(* IEC 61131-3 sources: Lasal-MCP/examples/SampleSource/LASALScreenAdvancedSolution/LASALScreenAdvancedSolution/LASALScreenAdvacnedSolution/Stations/Terminal/HMI/Class/MyRecalculate, 1 file *)

(* ---- MyRecalculate.st ---- *)
(*!
<Class
	Name               = "MyRecalculate"
	Revision           = "0.0"
	RealtimeTask       = "false"
	CyclicTask         = "false"
	BackgroundTask     = "false"
	Sigmatek           = "false"
	OSInterface        = "false"
	HighPriority       = "false"
	Automatic          = "false"
	UpdateMode         = "Prescan"
	SharedCommandTable = "true"
	Objectsize         = "(390,120)">
	<Channels>
		<Server Name="Length" Visualized="true" Initialize="false" WriteProtected="false" Retentive="false"/>
	</Channels>
	<Network Name="MyRecalculate">
		<!-- List of Components in this network -->
		<Components>
			<Object
				Name       = "_base"
				Class      = "_Global"
				Position   = "(218,120)"
				Visualized = "true"
				Remotely   = "true">
				<Channels>
					<Server Name="Server0"/>
					<Client Name="Lse"/>
				</Channels>
			</Object>
		</Components>
		<Comments>
		</Comments>
		<!-- List of Connections in this network -->
		<Connections>
			<Connection Source="this.Server0" Destination="_base.Server0" Vertices="(690,210),(518,210),"/>
			<Connection Source="_base.Lse" Destination="this.Lse" Vertices="(218,210),(38,210),"/>
		</Connections>
		<!-- Headerfiles -->
		<Options>
		</Options>
	</Network>
</Class>
*)
#pragma using _Global

MyRecalculate : CLASS
: _Global
  //Servers:
	Length 	: SvrCh_REAL;
  //Clients:
  //Variables:
  //Functions:
				//! <Function Comment="function is called in case of an recalculation (formula) defined for a data-server&#13;&#10;pres ....... --&gt; to value&#13;&#10;pv ......... --&gt; to variable&#13;&#10;direction .. direction (TRUE Y=kX+d, FALSE X=(Y+d)/k)&#13;&#10;retcode .... return TRUE if kernel should do the calculation, on the other hand return FALSE&#13;&#10;" Name="IF_Recalculate"/>
	FUNCTION VIRTUAL GLOBAL IF_Recalculate
		VAR_INPUT
			pres 	: ^_RESULT;
			pv 	: ^_VARIABLE;
			direction 	: BOOL;
		END_VAR
		VAR_OUTPUT
			retcode 	: BOOL;
		END_VAR;

	FUNCTION MeterToFeet
		VAR_INPUT
			value 	: REAL;
			dir 	: BOOL;
		END_VAR
		VAR_OUTPUT
			retcode 	: REAL;
		END_VAR;
  //Tables:
	FUNCTION @STD
		VAR_OUTPUT
			ret_code	: CONFSTATES;
		END_VAR;
	FUNCTION GLOBAL TAB @CT_;
END_CLASS;

FUNCTION VIRTUAL GLOBAL MyRecalculate::IF_Recalculate
	VAR_INPUT
		pres 	: ^_RESULT;
		pv 	: ^_VARIABLE;
		direction 	: BOOL;
	END_VAR
	VAR_OUTPUT
		retcode 	: BOOL;
	END_VAR

  retcode := TRUE;

  //====================================================================================
  case pv^.info.formula of

    //----------------------------------------------------------------------------------
    50: // The Formula number to be used for the unit

        pres^.value$REAL := MeterToFeet(value:= pres^.value$REAL, dir:= direction);

        retcode := FALSE;

  end_case;

END_FUNCTION

FUNCTION MyRecalculate::MeterToFeet
	VAR_INPUT
		value 	: REAL;
		dir 	: BOOL;
	END_VAR
	VAR_OUTPUT
		retcode 	: REAL;
	END_VAR

  if (dir = TRUE) then
    retCode := value / 0.3048;
  else
    retCode := value * 0.3048;
  end_if;

END_FUNCTION
